Fanuc KAREL source: KT00549.KL

PROGRAM KT00549
%NOLOCKGROUP
VAR
  P1: JOINTPOS
  P2: JOINTPOS
  OUT: POSITION
BEGIN
  OUT = P1 : P2
END KT00549
